Fanuc KAREL source: kt00343.KL

-- PROVISIONAL review KL for V770-1; original PC SHA256 24e771187fcb7b956ce496fdf9f39a0838c14bfb435fed8aaec904189a4fa9ec
-- Incomplete behavior may be omitted. Consult companion uncertainty JSON. Do not deploy.
PROGRAM KT00343
%NOLOCKGROUP
VAR
  I2 : INTEGER
  OUT : BOOLEAN
-- UNRESOLVED_DECL H1 type=002017
BEGIN
  -- UNRESOLVED_PC offsets 5-19; opcodes 2E,22,9D,33,B4
  -- UNRESOLVED_PC offsets 24-35; opcodes 2E,23
  -- UNRESOLVED_PC offsets 40-62; opcodes 22,9D,33,B3,21,59,23
  -- UNRESOLVED_PC offsets 67-71; opcodes 7F
END KT00343
